# EPICS substitutions: testIocApp/Db/BK9141.substitutions
file "$(TOP)/db/BK9141.db" {
  pattern
  { HWUNIT,   SYS,  SUB,  DEV,  INST    }
 { "BK9141",  "TST",  "", "PS", "N0001" }
}
